(* CoDeSys 2.3 export: ld.exp *)

(* POU PLC_LD_PRG_TR, LD *)
PROGRAM PLC_LD_PRG_TR
VAR
END_VAR
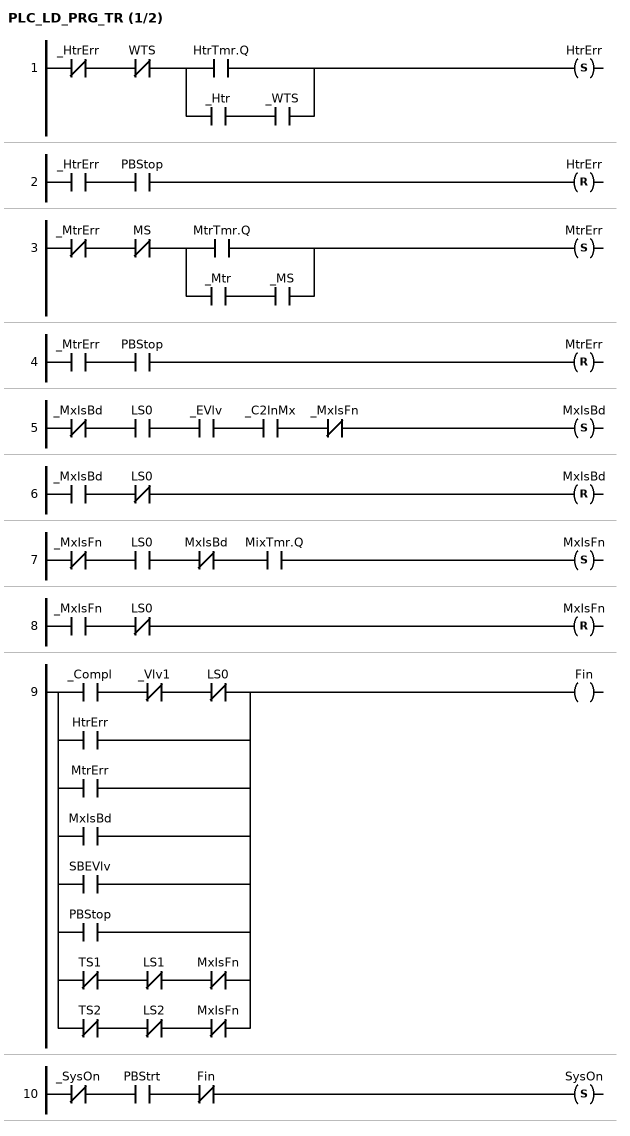
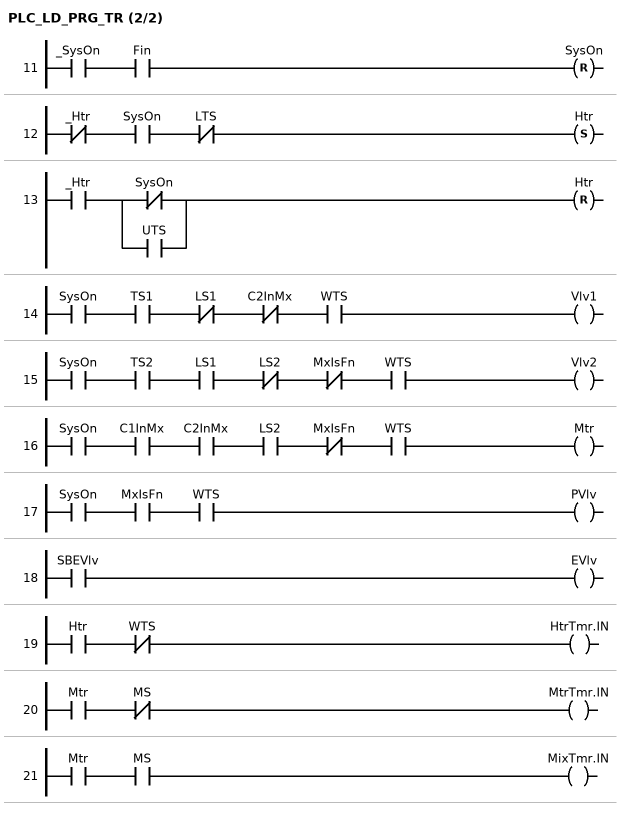
_LD_ (* Ladder Diagram *)
NETWORK 1
	[/_HtrErr] - [/WTS] - { [HtrTmr.Q] | [_Htr] - [_WTS] } --- (S HtrErr)
NETWORK 2
	[_HtrErr] - [PBStop] --- (R HtrErr)
NETWORK 3
	[/_MtrErr] - [/MS] - { [MtrTmr.Q] | [_Mtr] - [_MS] } --- (S MtrErr)
NETWORK 4
	[_MtrErr] - [PBStop] --- (R MtrErr)
NETWORK 5
	[/_MxIsBd] - [LS0] - [_EVlv] - [_C2InMx] - [/_MxIsFn] --- (S MxIsBd)
NETWORK 6
	[_MxIsBd] - [/LS0] --- (R MxIsBd)
NETWORK 7
	[/_MxIsFn] - [LS0] - [/MxIsBd] - [MixTmr.Q] --- (S MxIsFn)
NETWORK 8
	[_MxIsFn] - [/LS0] --- (R MxIsFn)
NETWORK 9
	{ [_Compl] - [/_Vlv1] - [/LS0] | [HtrErr] | [MtrErr] | [MxIsBd] | [SBEVlv] | [PBStop] | [/TS1] - [/LS1] - [/MxIsFn] | [/TS2] - [/LS2] - [/MxIsFn] } --- (Fin)
NETWORK 10
	[/_SysOn] - [PBStrt] - [/Fin] --- (S SysOn)
NETWORK 11
	[_SysOn] - [Fin] --- (R SysOn)
NETWORK 12
	[/_Htr] - [SysOn] - [/LTS] --- (S Htr)
NETWORK 13
	[_Htr] - { [/SysOn] | [UTS] } --- (R Htr)
NETWORK 14
	[SysOn] - [TS1] - [/LS1] - [/C2InMx] - [WTS] --- (Vlv1)
NETWORK 15
	[SysOn] - [TS2] - [LS1] - [/LS2] - [/MxIsFn] - [WTS] --- (Vlv2)
NETWORK 16
	[SysOn] - [C1InMx] - [C2InMx] - [LS2] - [/MxIsFn] - [WTS] --- (Mtr)
NETWORK 17
	[SysOn] - [MxIsFn] - [WTS] --- (PVlv)
NETWORK 18
	[SBEVlv] --- (EVlv)
NETWORK 19
	[Htr] - [/WTS] --- (HtrTmr.IN)
NETWORK 20
	[Mtr] - [/MS] --- (MtrTmr.IN)
NETWORK 21
	[Mtr] - [MS] --- (MixTmr.IN)
_END_LD_
(* the same logic as Structured Text *)
(* Network 1 *)
IF NOT _HtrErr AND NOT WTS AND (HtrTmr.Q OR _Htr AND _WTS) THEN HtrErr := TRUE; END_IF;
(* Network 2 *)
IF _HtrErr AND PBStop THEN HtrErr := FALSE; END_IF;
(* Network 3 *)
IF NOT _MtrErr AND NOT MS AND (MtrTmr.Q OR _Mtr AND _MS) THEN MtrErr := TRUE; END_IF;
(* Network 4 *)
IF _MtrErr AND PBStop THEN MtrErr := FALSE; END_IF;
(* Network 5 *)
IF NOT _MxIsBd AND LS0 AND _EVlv AND _C2InMx AND NOT _MxIsFn THEN MxIsBd := TRUE; END_IF;
(* Network 6 *)
IF _MxIsBd AND NOT LS0 THEN MxIsBd := FALSE; END_IF;
(* Network 7 *)
IF NOT _MxIsFn AND LS0 AND NOT MxIsBd AND MixTmr.Q THEN MxIsFn := TRUE; END_IF;
(* Network 8 *)
IF _MxIsFn AND NOT LS0 THEN MxIsFn := FALSE; END_IF;
(* Network 9 *)
Fin := _Compl AND NOT _Vlv1 AND NOT LS0 OR HtrErr OR MtrErr OR MxIsBd OR SBEVlv OR PBStop OR NOT TS1 AND NOT LS1 AND NOT MxIsFn OR NOT TS2 AND NOT LS2 AND NOT MxIsFn;
(* Network 10 *)
IF NOT _SysOn AND PBStrt AND NOT Fin THEN SysOn := TRUE; END_IF;
(* Network 11 *)
IF _SysOn AND Fin THEN SysOn := FALSE; END_IF;
(* Network 12 *)
IF NOT _Htr AND SysOn AND NOT LTS THEN Htr := TRUE; END_IF;
(* Network 13 *)
IF _Htr AND (NOT SysOn OR UTS) THEN Htr := FALSE; END_IF;
(* Network 14 *)
Vlv1 := SysOn AND TS1 AND NOT LS1 AND NOT C2InMx AND WTS;
(* Network 15 *)
Vlv2 := SysOn AND TS2 AND LS1 AND NOT LS2 AND NOT MxIsFn AND WTS;
(* Network 16 *)
Mtr := SysOn AND C1InMx AND C2InMx AND LS2 AND NOT MxIsFn AND WTS;
(* Network 17 *)
PVlv := SysOn AND MxIsFn AND WTS;
(* Network 18 *)
EVlv := SBEVlv;
(* Network 19 *)
HtrTmr.IN := Htr AND NOT WTS;
(* Network 20 *)
MtrTmr.IN := Mtr AND NOT MS;
(* Network 21 *)
MixTmr.IN := Mtr AND MS;
END_PROGRAM
